(* IEC 61131-3 sources: nautilus/examples/plclab, 2 files *)

(* ---- types.st ---- *)
(* The connector PLC-Lab reads and writes over OPC UA. PLC-Lab looks for a
   container named exactly PlcLabConnector holding these members, with these
   names and types: on CODESYS it is a global variable list; here it is one
   struct tag of this type (nautilus.yaml). See README.md.

   PLC-Lab writes Inputs (its sensors, as bytes) and the two area tables,
   which say which bytes it uses; it reads Outputs. The SIZE_ members tell it
   how big the arrays are. *)

TYPE
  PlcLabArea : STRUCT
    CntBytes : WORD;  (* how many bytes; 0 ends the table *)
    Addr     : WORD;  (* first byte in Inputs or Outputs *)
    IoOfs    : WORD;  (* first byte of the process image: 0 is IB0 / QB0 *)
  END_STRUCT;

  PlcLabConnectorData : STRUCT
    SIZE_AREA_I_ARRAY : WORD := 10;
    SIZE_AREA_Q_ARRAY : WORD := 10;
    SIZE_I_ARRAY      : WORD := 1024;
    SIZE_Q_ARRAY      : WORD := 1024;
    Inputs      : ARRAY[0..1023] OF BYTE;      (* written by PLC-Lab *)
    Outputs     : ARRAY[0..1023] OF BYTE;      (* read by PLC-Lab *)
    AreaInputs  : ARRAY[0..9] OF PlcLabArea;   (* written by PLC-Lab *)
    AreaOutputs : ARRAY[0..9] OF PlcLabArea;   (* written by PLC-Lab *)
  END_STRUCT;
END_TYPE

(* ---- plclab.st ---- *)
PROGRAM PlcLab
(* One scan: PLC-Lab's input bytes into the process image, the image's
   bits onto named tags, the tank logic, and the outputs back into the bytes
   PLC-Lab reads. The connector half is what PlcLabSync does on CODESYS,
   written without pointers: the process image is two local byte arrays,
   IB0..IB15 and QB0..QB15, and a sensor PLC-Lab calls I0.2 is bit 2 of
   ib[0].

   The area tables say where things are. Area a copies CntBytes bytes:
   Inputs[Addr + i] into ib[IoOfs + i], and qb[IoOfs + i] into
   Outputs[Addr + i]. The first area with CntBytes = 0 ends the table. A
   byte outside the connector or the image is skipped, never a fault. *)
VAR_EXTERNAL
    PlcLabConnector : PlcLabConnectorData;
    PlcLabMapped : BOOL;

    StartPB   : BOOL;
    StopPB    : BOOL;
    LevelLow  : BOOL;
    LevelHigh : BOOL;

    FillValve  : BOOL;
    DrainValve : BOOL;
    RunLamp    : BOOL;
    FullLamp   : BOOL;
END_VAR
VAR
    ib : ARRAY[0..15] OF BYTE;  (* inputs as PLC-Lab numbers them: ib[0] is IB0 *)
    qb : ARRAY[0..15] OF BYTE;  (* outputs: qb[0] is QB0 *)
    a, i, n, src, dst : DINT;
    tank : TankCycle;
END_VAR

(* PLC-Lab's input bytes into the image *)
FOR a := 0 TO 9 DO
    n := PlcLabConnector.AreaInputs[a].CntBytes;
    IF n = 0 THEN
        EXIT;
    END_IF;
    FOR i := 0 TO n - 1 DO
        src := PlcLabConnector.AreaInputs[a].Addr + i;
        dst := PlcLabConnector.AreaInputs[a].IoOfs + i;
        IF src <= 1023 AND dst <= 15 THEN
            ib[dst] := PlcLabConnector.Inputs[src];
        END_IF;
    END_FOR;
END_FOR;
PlcLabMapped := PlcLabConnector.AreaInputs[0].CntBytes > 0 OR PlcLabConnector.AreaOutputs[0].CntBytes > 0;

(* the image's bits onto named tags *)
StartPB   := ib[0].%X0;  (* I0.0 *)
StopPB    := ib[0].%X1;  (* I0.1, normally closed *)
LevelLow  := ib[0].%X2;  (* I0.2 *)
LevelHigh := ib[0].%X3;  (* I0.3 *)

tank(Start := StartPB, Stop := StopPB, Low := LevelLow, High := LevelHigh);
FillValve  := tank.Fill;
DrainValve := tank.Drain;
RunLamp    := tank.Running;
FullLamp   := tank.Full;

qb[0].%X0 := FillValve;   (* Q0.0 *)
qb[0].%X1 := DrainValve;  (* Q0.1 *)
qb[0].%X2 := RunLamp;     (* Q0.2 *)
qb[0].%X3 := FullLamp;    (* Q0.3 *)

(* the image into the bytes PLC-Lab reads. The commit at the end of the
   scan lands only the Outputs bytes assigned here, so an input byte or an
   area entry PLC-Lab writes while the scan runs is never put back. *)
FOR a := 0 TO 9 DO
    n := PlcLabConnector.AreaOutputs[a].CntBytes;
    IF n = 0 THEN
        EXIT;
    END_IF;
    FOR i := 0 TO n - 1 DO
        src := PlcLabConnector.AreaOutputs[a].IoOfs + i;
        dst := PlcLabConnector.AreaOutputs[a].Addr + i;
        IF src <= 15 AND dst <= 1023 THEN
            PlcLabConnector.Outputs[dst] := qb[src];
        END_IF;
    END_FOR;
END_FOR;
END_PROGRAM
